FUNCTION "FRK_LineSetWalk" : Bool
{ S7_Optimized_Access := 'TRUE' }
VERSION : 0.1
VAR_INPUT
    RootIndex : Int;
    Scope : String;
    Phase : Int;
    Access : "FRK_Access";
    Ready : Bool;
END_VAR
VAR_TEMP
    Slot : Int;
END_VAR
BEGIN
    #FRK_LineSetWalk := FALSE;
    "FRK_SetRuntime".Work[#RootIndex].RejectScope := 'BenchLineOwner';
    IF NOT "FRK_LineScope"(Scope := #Scope) OR NOT "FRK_Line".Data.Applied
        OR "FRK_Line".Data.Status.Role <> 1 THEN RETURN; END_IF;
    IF #Phase = 2 THEN
        "FRK_Line".Data.Values := "FRK_LineSetStage".Values;
        "FRK_LineCommit"(State := "FRK_Line".Data);
        #FRK_LineSetWalk := TRUE; RETURN;
    END_IF;
    IF #Phase = 1 OR #Phase = 4 THEN "FRK_LineSetStage".Values := "FRK_Line".Data.Values; END_IF;
    "FRK_LineDef"(FieldIndex := 1);
    "FRK_SetRuntime".Work[#RootIndex].RejectScope := #Scope; "FRK_SetRuntime".Work[#RootIndex].RejectKey := "FRK_ConfigScratch".Entry.WriteKey;
    IF #Phase = 0 OR #Phase = 5 THEN
        IF #Phase = 5 AND NOT "FRK_ConfigDataAllowed"(Access := #Access, ForWrite := FALSE, Scope := #Scope) THEN RETURN; END_IF;
        "FRK_LineValue"(FieldIndex := 1, Values := "FRK_Line".Data.Values);
        IF NOT "FRK_ConfigValidate"(Text := "FRK_ConfigScratch".Entry.ValueText)
            OR "FRK_SetRuntime".Work[#RootIndex].Payload.Info.RecordCount >= 29 THEN RETURN; END_IF;
        #Slot := "FRK_SetRuntime".Work[#RootIndex].Payload.Info.RecordCount + 1;
        "FRK_SetRuntime".Work[#RootIndex].Payload.Records[#Slot].Scope := #Scope;
        "FRK_SetRuntime".Work[#RootIndex].Payload.Records[#Slot].WriteKey := "FRK_ConfigScratch".Entry.WriteKey;
        "FRK_SetRuntime".Work[#RootIndex].Payload.Records[#Slot].Revision := "FRK_ConfigScratch".Entry.WriteRevision;
        "FRK_SetRuntime".Work[#RootIndex].Payload.Records[#Slot].Kind := "FRK_ConfigScratch".Entry.ConfigKind;
        "FRK_SetRuntime".Work[#RootIndex].Payload.Records[#Slot].ValueType := "FRK_ConfigScratch".Entry.ValueType;
        "FRK_SetRuntime".Work[#RootIndex].Payload.Records[#Slot].ValueText := WSTRING_TO_STRING("FRK_ConfigScratch".Entry.ValueText);
        "FRK_SetRuntime".Work[#RootIndex].Payload.Info.RecordCount := #Slot;
    ELSE
        #Slot := "FRK_SetCheck"(RootIndex := #RootIndex, Scope := #Scope, Access := #Access, Ready := #Ready AND (#Phase = 4 OR "FRK_Line".Ready), WriteAccess := #Phase <> 3, ReserveTarget := FALSE);
        IF #Slot = 0 THEN RETURN; END_IF;
        IF #Phase = 1 OR #Phase = 4 THEN
    "FRK_LineSetStage".Values.TaktMs := LINT_TO_UDINT("FRK_ConfigScratch".Value.Number);
        END_IF;
    END_IF;
    "FRK_LineDef"(FieldIndex := 2);
    "FRK_SetRuntime".Work[#RootIndex].RejectScope := #Scope; "FRK_SetRuntime".Work[#RootIndex].RejectKey := "FRK_ConfigScratch".Entry.WriteKey;
    IF #Phase = 0 OR #Phase = 5 THEN
        IF #Phase = 5 AND NOT "FRK_ConfigDataAllowed"(Access := #Access, ForWrite := FALSE, Scope := #Scope) THEN RETURN; END_IF;
        "FRK_LineValue"(FieldIndex := 2, Values := "FRK_Line".Data.Values);
        IF NOT "FRK_ConfigValidate"(Text := "FRK_ConfigScratch".Entry.ValueText)
            OR "FRK_SetRuntime".Work[#RootIndex].Payload.Info.RecordCount >= 29 THEN RETURN; END_IF;
        #Slot := "FRK_SetRuntime".Work[#RootIndex].Payload.Info.RecordCount + 1;
        "FRK_SetRuntime".Work[#RootIndex].Payload.Records[#Slot].Scope := #Scope;
        "FRK_SetRuntime".Work[#RootIndex].Payload.Records[#Slot].WriteKey := "FRK_ConfigScratch".Entry.WriteKey;
        "FRK_SetRuntime".Work[#RootIndex].Payload.Records[#Slot].Revision := "FRK_ConfigScratch".Entry.WriteRevision;
        "FRK_SetRuntime".Work[#RootIndex].Payload.Records[#Slot].Kind := "FRK_ConfigScratch".Entry.ConfigKind;
        "FRK_SetRuntime".Work[#RootIndex].Payload.Records[#Slot].ValueType := "FRK_ConfigScratch".Entry.ValueType;
        "FRK_SetRuntime".Work[#RootIndex].Payload.Records[#Slot].ValueText := WSTRING_TO_STRING("FRK_ConfigScratch".Entry.ValueText);
        "FRK_SetRuntime".Work[#RootIndex].Payload.Info.RecordCount := #Slot;
    ELSE
        #Slot := "FRK_SetCheck"(RootIndex := #RootIndex, Scope := #Scope, Access := #Access, Ready := #Ready AND (#Phase = 4 OR "FRK_Line".Ready), WriteAccess := #Phase <> 3, ReserveTarget := FALSE);
        IF #Slot = 0 THEN RETURN; END_IF;
        IF #Phase = 1 OR #Phase = 4 THEN
    "FRK_LineSetStage".Values.Gain := "FRK_ConfigScratch".Value.Decimal;
        END_IF;
    END_IF;
    "FRK_LineDef"(FieldIndex := 3);
    "FRK_SetRuntime".Work[#RootIndex].RejectScope := #Scope; "FRK_SetRuntime".Work[#RootIndex].RejectKey := "FRK_ConfigScratch".Entry.WriteKey;
    IF #Phase = 0 OR #Phase = 5 THEN
        IF #Phase = 5 AND NOT "FRK_ConfigDataAllowed"(Access := #Access, ForWrite := FALSE, Scope := #Scope) THEN RETURN; END_IF;
        "FRK_LineValue"(FieldIndex := 3, Values := "FRK_Line".Data.Values);
        IF NOT "FRK_ConfigValidate"(Text := "FRK_ConfigScratch".Entry.ValueText)
            OR "FRK_SetRuntime".Work[#RootIndex].Payload.Info.RecordCount >= 29 THEN RETURN; END_IF;
        #Slot := "FRK_SetRuntime".Work[#RootIndex].Payload.Info.RecordCount + 1;
        "FRK_SetRuntime".Work[#RootIndex].Payload.Records[#Slot].Scope := #Scope;
        "FRK_SetRuntime".Work[#RootIndex].Payload.Records[#Slot].WriteKey := "FRK_ConfigScratch".Entry.WriteKey;
        "FRK_SetRuntime".Work[#RootIndex].Payload.Records[#Slot].Revision := "FRK_ConfigScratch".Entry.WriteRevision;
        "FRK_SetRuntime".Work[#RootIndex].Payload.Records[#Slot].Kind := "FRK_ConfigScratch".Entry.ConfigKind;
        "FRK_SetRuntime".Work[#RootIndex].Payload.Records[#Slot].ValueType := "FRK_ConfigScratch".Entry.ValueType;
        "FRK_SetRuntime".Work[#RootIndex].Payload.Records[#Slot].ValueText := WSTRING_TO_STRING("FRK_ConfigScratch".Entry.ValueText);
        "FRK_SetRuntime".Work[#RootIndex].Payload.Info.RecordCount := #Slot;
    ELSE
        #Slot := "FRK_SetCheck"(RootIndex := #RootIndex, Scope := #Scope, Access := #Access, Ready := #Ready AND (#Phase = 4 OR "FRK_Line".Ready), WriteAccess := #Phase <> 3, ReserveTarget := FALSE);
        IF #Slot = 0 THEN RETURN; END_IF;
        IF #Phase = 1 OR #Phase = 4 THEN
    "FRK_LineSetStage".Values.Grade := LINT_TO_DINT("FRK_ConfigScratch".Value.Number);
        END_IF;
    END_IF;
    "FRK_LineDef"(FieldIndex := 4);
    "FRK_SetRuntime".Work[#RootIndex].RejectScope := #Scope; "FRK_SetRuntime".Work[#RootIndex].RejectKey := "FRK_ConfigScratch".Entry.WriteKey;
    IF #Phase = 0 OR #Phase = 5 THEN
        IF #Phase = 5 AND NOT "FRK_ConfigDataAllowed"(Access := #Access, ForWrite := FALSE, Scope := #Scope) THEN RETURN; END_IF;
        "FRK_LineValue"(FieldIndex := 4, Values := "FRK_Line".Data.Values);
        IF NOT "FRK_ConfigValidate"(Text := "FRK_ConfigScratch".Entry.ValueText)
            OR "FRK_SetRuntime".Work[#RootIndex].Payload.Info.RecordCount >= 29 THEN RETURN; END_IF;
        #Slot := "FRK_SetRuntime".Work[#RootIndex].Payload.Info.RecordCount + 1;
        "FRK_SetRuntime".Work[#RootIndex].Payload.Records[#Slot].Scope := #Scope;
        "FRK_SetRuntime".Work[#RootIndex].Payload.Records[#Slot].WriteKey := "FRK_ConfigScratch".Entry.WriteKey;
        "FRK_SetRuntime".Work[#RootIndex].Payload.Records[#Slot].Revision := "FRK_ConfigScratch".Entry.WriteRevision;
        "FRK_SetRuntime".Work[#RootIndex].Payload.Records[#Slot].Kind := "FRK_ConfigScratch".Entry.ConfigKind;
        "FRK_SetRuntime".Work[#RootIndex].Payload.Records[#Slot].ValueType := "FRK_ConfigScratch".Entry.ValueType;
        "FRK_SetRuntime".Work[#RootIndex].Payload.Records[#Slot].ValueText := WSTRING_TO_STRING("FRK_ConfigScratch".Entry.ValueText);
        "FRK_SetRuntime".Work[#RootIndex].Payload.Info.RecordCount := #Slot;
    ELSE
        #Slot := "FRK_SetCheck"(RootIndex := #RootIndex, Scope := #Scope, Access := #Access, Ready := #Ready AND (#Phase = 4 OR "FRK_Line".Ready), WriteAccess := #Phase <> 3, ReserveTarget := FALSE);
        IF #Slot = 0 THEN RETURN; END_IF;
        IF #Phase = 1 OR #Phase = 4 THEN
    "FRK_LineSetStage".Values.Enabled := "FRK_ConfigScratch".Value.Flag;
        END_IF;
    END_IF;
    "FRK_LineDef"(FieldIndex := 5);
    "FRK_SetRuntime".Work[#RootIndex].RejectScope := #Scope; "FRK_SetRuntime".Work[#RootIndex].RejectKey := "FRK_ConfigScratch".Entry.WriteKey;
    IF #Phase = 0 OR #Phase = 5 THEN
        IF #Phase = 5 AND NOT "FRK_ConfigDataAllowed"(Access := #Access, ForWrite := FALSE, Scope := #Scope) THEN RETURN; END_IF;
        "FRK_LineValue"(FieldIndex := 5, Values := "FRK_Line".Data.Values);
        IF NOT "FRK_ConfigValidate"(Text := "FRK_ConfigScratch".Entry.ValueText)
            OR "FRK_SetRuntime".Work[#RootIndex].Payload.Info.RecordCount >= 29 THEN RETURN; END_IF;
        #Slot := "FRK_SetRuntime".Work[#RootIndex].Payload.Info.RecordCount + 1;
        "FRK_SetRuntime".Work[#RootIndex].Payload.Records[#Slot].Scope := #Scope;
        "FRK_SetRuntime".Work[#RootIndex].Payload.Records[#Slot].WriteKey := "FRK_ConfigScratch".Entry.WriteKey;
        "FRK_SetRuntime".Work[#RootIndex].Payload.Records[#Slot].Revision := "FRK_ConfigScratch".Entry.WriteRevision;
        "FRK_SetRuntime".Work[#RootIndex].Payload.Records[#Slot].Kind := "FRK_ConfigScratch".Entry.ConfigKind;
        "FRK_SetRuntime".Work[#RootIndex].Payload.Records[#Slot].ValueType := "FRK_ConfigScratch".Entry.ValueType;
        "FRK_SetRuntime".Work[#RootIndex].Payload.Records[#Slot].ValueText := WSTRING_TO_STRING("FRK_ConfigScratch".Entry.ValueText);
        "FRK_SetRuntime".Work[#RootIndex].Payload.Info.RecordCount := #Slot;
    ELSE
        #Slot := "FRK_SetCheck"(RootIndex := #RootIndex, Scope := #Scope, Access := #Access, Ready := #Ready AND (#Phase = 4 OR "FRK_Line".Ready), WriteAccess := #Phase <> 3, ReserveTarget := FALSE);
        IF #Slot = 0 THEN RETURN; END_IF;
        IF #Phase = 1 OR #Phase = 4 THEN
    "FRK_LineSetStage".Values.HostName := "FRK_ConfigScratch".Value.Text;
        END_IF;
    END_IF;
    "FRK_LineDef"(FieldIndex := 6);
    "FRK_SetRuntime".Work[#RootIndex].RejectScope := #Scope; "FRK_SetRuntime".Work[#RootIndex].RejectKey := "FRK_ConfigScratch".Entry.WriteKey;
    IF #Phase = 0 OR #Phase = 5 THEN
        IF #Phase = 5 AND NOT "FRK_ConfigDataAllowed"(Access := #Access, ForWrite := FALSE, Scope := #Scope) THEN RETURN; END_IF;
        "FRK_LineValue"(FieldIndex := 6, Values := "FRK_Line".Data.Values);
        IF NOT "FRK_ConfigValidate"(Text := "FRK_ConfigScratch".Entry.ValueText)
            OR "FRK_SetRuntime".Work[#RootIndex].Payload.Info.RecordCount >= 29 THEN RETURN; END_IF;
        #Slot := "FRK_SetRuntime".Work[#RootIndex].Payload.Info.RecordCount + 1;
        "FRK_SetRuntime".Work[#RootIndex].Payload.Records[#Slot].Scope := #Scope;
        "FRK_SetRuntime".Work[#RootIndex].Payload.Records[#Slot].WriteKey := "FRK_ConfigScratch".Entry.WriteKey;
        "FRK_SetRuntime".Work[#RootIndex].Payload.Records[#Slot].Revision := "FRK_ConfigScratch".Entry.WriteRevision;
        "FRK_SetRuntime".Work[#RootIndex].Payload.Records[#Slot].Kind := "FRK_ConfigScratch".Entry.ConfigKind;
        "FRK_SetRuntime".Work[#RootIndex].Payload.Records[#Slot].ValueType := "FRK_ConfigScratch".Entry.ValueType;
        "FRK_SetRuntime".Work[#RootIndex].Payload.Records[#Slot].ValueText := WSTRING_TO_STRING("FRK_ConfigScratch".Entry.ValueText);
        "FRK_SetRuntime".Work[#RootIndex].Payload.Info.RecordCount := #Slot;
    ELSE
        #Slot := "FRK_SetCheck"(RootIndex := #RootIndex, Scope := #Scope, Access := #Access, Ready := #Ready AND (#Phase = 4 OR "FRK_Line".Ready), WriteAccess := #Phase <> 3, ReserveTarget := FALSE);
        IF #Slot = 0 THEN RETURN; END_IF;
        IF #Phase = 1 OR #Phase = 4 THEN
    "FRK_LineSetStage".Values.Offsets[0] := LINT_TO_INT("FRK_ConfigScratch".Value.Number);
        END_IF;
    END_IF;
    "FRK_LineDef"(FieldIndex := 7);
    "FRK_SetRuntime".Work[#RootIndex].RejectScope := #Scope; "FRK_SetRuntime".Work[#RootIndex].RejectKey := "FRK_ConfigScratch".Entry.WriteKey;
    IF #Phase = 0 OR #Phase = 5 THEN
        IF #Phase = 5 AND NOT "FRK_ConfigDataAllowed"(Access := #Access, ForWrite := FALSE, Scope := #Scope) THEN RETURN; END_IF;
        "FRK_LineValue"(FieldIndex := 7, Values := "FRK_Line".Data.Values);
        IF NOT "FRK_ConfigValidate"(Text := "FRK_ConfigScratch".Entry.ValueText)
            OR "FRK_SetRuntime".Work[#RootIndex].Payload.Info.RecordCount >= 29 THEN RETURN; END_IF;
        #Slot := "FRK_SetRuntime".Work[#RootIndex].Payload.Info.RecordCount + 1;
        "FRK_SetRuntime".Work[#RootIndex].Payload.Records[#Slot].Scope := #Scope;
        "FRK_SetRuntime".Work[#RootIndex].Payload.Records[#Slot].WriteKey := "FRK_ConfigScratch".Entry.WriteKey;
        "FRK_SetRuntime".Work[#RootIndex].Payload.Records[#Slot].Revision := "FRK_ConfigScratch".Entry.WriteRevision;
        "FRK_SetRuntime".Work[#RootIndex].Payload.Records[#Slot].Kind := "FRK_ConfigScratch".Entry.ConfigKind;
        "FRK_SetRuntime".Work[#RootIndex].Payload.Records[#Slot].ValueType := "FRK_ConfigScratch".Entry.ValueType;
        "FRK_SetRuntime".Work[#RootIndex].Payload.Records[#Slot].ValueText := WSTRING_TO_STRING("FRK_ConfigScratch".Entry.ValueText);
        "FRK_SetRuntime".Work[#RootIndex].Payload.Info.RecordCount := #Slot;
    ELSE
        #Slot := "FRK_SetCheck"(RootIndex := #RootIndex, Scope := #Scope, Access := #Access, Ready := #Ready AND (#Phase = 4 OR "FRK_Line".Ready), WriteAccess := #Phase <> 3, ReserveTarget := FALSE);
        IF #Slot = 0 THEN RETURN; END_IF;
        IF #Phase = 1 OR #Phase = 4 THEN
    "FRK_LineSetStage".Values.Offsets[1] := LINT_TO_INT("FRK_ConfigScratch".Value.Number);
        END_IF;
    END_IF;
    "FRK_LineDef"(FieldIndex := 8);
    "FRK_SetRuntime".Work[#RootIndex].RejectScope := #Scope; "FRK_SetRuntime".Work[#RootIndex].RejectKey := "FRK_ConfigScratch".Entry.WriteKey;
    IF #Phase = 0 OR #Phase = 5 THEN
        IF #Phase = 5 AND NOT "FRK_ConfigDataAllowed"(Access := #Access, ForWrite := FALSE, Scope := #Scope) THEN RETURN; END_IF;
        "FRK_LineValue"(FieldIndex := 8, Values := "FRK_Line".Data.Values);
        IF NOT "FRK_ConfigValidate"(Text := "FRK_ConfigScratch".Entry.ValueText)
            OR "FRK_SetRuntime".Work[#RootIndex].Payload.Info.RecordCount >= 29 THEN RETURN; END_IF;
        #Slot := "FRK_SetRuntime".Work[#RootIndex].Payload.Info.RecordCount + 1;
        "FRK_SetRuntime".Work[#RootIndex].Payload.Records[#Slot].Scope := #Scope;
        "FRK_SetRuntime".Work[#RootIndex].Payload.Records[#Slot].WriteKey := "FRK_ConfigScratch".Entry.WriteKey;
        "FRK_SetRuntime".Work[#RootIndex].Payload.Records[#Slot].Revision := "FRK_ConfigScratch".Entry.WriteRevision;
        "FRK_SetRuntime".Work[#RootIndex].Payload.Records[#Slot].Kind := "FRK_ConfigScratch".Entry.ConfigKind;
        "FRK_SetRuntime".Work[#RootIndex].Payload.Records[#Slot].ValueType := "FRK_ConfigScratch".Entry.ValueType;
        "FRK_SetRuntime".Work[#RootIndex].Payload.Records[#Slot].ValueText := WSTRING_TO_STRING("FRK_ConfigScratch".Entry.ValueText);
        "FRK_SetRuntime".Work[#RootIndex].Payload.Info.RecordCount := #Slot;
    ELSE
        #Slot := "FRK_SetCheck"(RootIndex := #RootIndex, Scope := #Scope, Access := #Access, Ready := #Ready AND (#Phase = 4 OR "FRK_Line".Ready), WriteAccess := #Phase <> 3, ReserveTarget := FALSE);
        IF #Slot = 0 THEN RETURN; END_IF;
        IF #Phase = 1 OR #Phase = 4 THEN
    "FRK_LineSetStage".Values.Small := LINT_TO_USINT("FRK_ConfigScratch".Value.Number);
        END_IF;
    END_IF;
    "FRK_LineDef"(FieldIndex := 9);
    "FRK_SetRuntime".Work[#RootIndex].RejectScope := #Scope; "FRK_SetRuntime".Work[#RootIndex].RejectKey := "FRK_ConfigScratch".Entry.WriteKey;
    IF #Phase = 0 OR #Phase = 5 THEN
        IF #Phase = 5 AND NOT "FRK_ConfigDataAllowed"(Access := #Access, ForWrite := FALSE, Scope := #Scope) THEN RETURN; END_IF;
        "FRK_LineValue"(FieldIndex := 9, Values := "FRK_Line".Data.Values);
        IF NOT "FRK_ConfigValidate"(Text := "FRK_ConfigScratch".Entry.ValueText)
            OR "FRK_SetRuntime".Work[#RootIndex].Payload.Info.RecordCount >= 29 THEN RETURN; END_IF;
        #Slot := "FRK_SetRuntime".Work[#RootIndex].Payload.Info.RecordCount + 1;
        "FRK_SetRuntime".Work[#RootIndex].Payload.Records[#Slot].Scope := #Scope;
        "FRK_SetRuntime".Work[#RootIndex].Payload.Records[#Slot].WriteKey := "FRK_ConfigScratch".Entry.WriteKey;
        "FRK_SetRuntime".Work[#RootIndex].Payload.Records[#Slot].Revision := "FRK_ConfigScratch".Entry.WriteRevision;
        "FRK_SetRuntime".Work[#RootIndex].Payload.Records[#Slot].Kind := "FRK_ConfigScratch".Entry.ConfigKind;
        "FRK_SetRuntime".Work[#RootIndex].Payload.Records[#Slot].ValueType := "FRK_ConfigScratch".Entry.ValueType;
        "FRK_SetRuntime".Work[#RootIndex].Payload.Records[#Slot].ValueText := WSTRING_TO_STRING("FRK_ConfigScratch".Entry.ValueText);
        "FRK_SetRuntime".Work[#RootIndex].Payload.Info.RecordCount := #Slot;
    ELSE
        #Slot := "FRK_SetCheck"(RootIndex := #RootIndex, Scope := #Scope, Access := #Access, Ready := #Ready AND (#Phase = 4 OR "FRK_Line".Ready), WriteAccess := #Phase <> 3, ReserveTarget := FALSE);
        IF #Slot = 0 THEN RETURN; END_IF;
        IF #Phase = 1 OR #Phase = 4 THEN
    "FRK_LineSetStage".Values.UtcOffsetMin := LINT_TO_DINT("FRK_ConfigScratch".Value.Number);
        END_IF;
    END_IF;
    "FRK_LineDef"(FieldIndex := 10);
    "FRK_SetRuntime".Work[#RootIndex].RejectScope := #Scope; "FRK_SetRuntime".Work[#RootIndex].RejectKey := "FRK_ConfigScratch".Entry.WriteKey;
    IF #Phase = 0 OR #Phase = 5 THEN
        IF #Phase = 5 AND NOT "FRK_ConfigDataAllowed"(Access := #Access, ForWrite := FALSE, Scope := #Scope) THEN RETURN; END_IF;
        "FRK_LineValue"(FieldIndex := 10, Values := "FRK_Line".Data.Values);
        IF NOT "FRK_ConfigValidate"(Text := "FRK_ConfigScratch".Entry.ValueText)
            OR "FRK_SetRuntime".Work[#RootIndex].Payload.Info.RecordCount >= 29 THEN RETURN; END_IF;
        #Slot := "FRK_SetRuntime".Work[#RootIndex].Payload.Info.RecordCount + 1;
        "FRK_SetRuntime".Work[#RootIndex].Payload.Records[#Slot].Scope := #Scope;
        "FRK_SetRuntime".Work[#RootIndex].Payload.Records[#Slot].WriteKey := "FRK_ConfigScratch".Entry.WriteKey;
        "FRK_SetRuntime".Work[#RootIndex].Payload.Records[#Slot].Revision := "FRK_ConfigScratch".Entry.WriteRevision;
        "FRK_SetRuntime".Work[#RootIndex].Payload.Records[#Slot].Kind := "FRK_ConfigScratch".Entry.ConfigKind;
        "FRK_SetRuntime".Work[#RootIndex].Payload.Records[#Slot].ValueType := "FRK_ConfigScratch".Entry.ValueType;
        "FRK_SetRuntime".Work[#RootIndex].Payload.Records[#Slot].ValueText := WSTRING_TO_STRING("FRK_ConfigScratch".Entry.ValueText);
        "FRK_SetRuntime".Work[#RootIndex].Payload.Info.RecordCount := #Slot;
    ELSE
        #Slot := "FRK_SetCheck"(RootIndex := #RootIndex, Scope := #Scope, Access := #Access, Ready := #Ready AND (#Phase = 4 OR "FRK_Line".Ready), WriteAccess := #Phase <> 3, ReserveTarget := FALSE);
        IF #Slot = 0 THEN RETURN; END_IF;
        IF #Phase = 1 OR #Phase = 4 THEN
    "FRK_LineSetStage".Values.ShiftStartMin[1] := LINT_TO_DINT("FRK_ConfigScratch".Value.Number);
        END_IF;
    END_IF;
    "FRK_LineDef"(FieldIndex := 11);
    "FRK_SetRuntime".Work[#RootIndex].RejectScope := #Scope; "FRK_SetRuntime".Work[#RootIndex].RejectKey := "FRK_ConfigScratch".Entry.WriteKey;
    IF #Phase = 0 OR #Phase = 5 THEN
        IF #Phase = 5 AND NOT "FRK_ConfigDataAllowed"(Access := #Access, ForWrite := FALSE, Scope := #Scope) THEN RETURN; END_IF;
        "FRK_LineValue"(FieldIndex := 11, Values := "FRK_Line".Data.Values);
        IF NOT "FRK_ConfigValidate"(Text := "FRK_ConfigScratch".Entry.ValueText)
            OR "FRK_SetRuntime".Work[#RootIndex].Payload.Info.RecordCount >= 29 THEN RETURN; END_IF;
        #Slot := "FRK_SetRuntime".Work[#RootIndex].Payload.Info.RecordCount + 1;
        "FRK_SetRuntime".Work[#RootIndex].Payload.Records[#Slot].Scope := #Scope;
        "FRK_SetRuntime".Work[#RootIndex].Payload.Records[#Slot].WriteKey := "FRK_ConfigScratch".Entry.WriteKey;
        "FRK_SetRuntime".Work[#RootIndex].Payload.Records[#Slot].Revision := "FRK_ConfigScratch".Entry.WriteRevision;
        "FRK_SetRuntime".Work[#RootIndex].Payload.Records[#Slot].Kind := "FRK_ConfigScratch".Entry.ConfigKind;
        "FRK_SetRuntime".Work[#RootIndex].Payload.Records[#Slot].ValueType := "FRK_ConfigScratch".Entry.ValueType;
        "FRK_SetRuntime".Work[#RootIndex].Payload.Records[#Slot].ValueText := WSTRING_TO_STRING("FRK_ConfigScratch".Entry.ValueText);
        "FRK_SetRuntime".Work[#RootIndex].Payload.Info.RecordCount := #Slot;
    ELSE
        #Slot := "FRK_SetCheck"(RootIndex := #RootIndex, Scope := #Scope, Access := #Access, Ready := #Ready AND (#Phase = 4 OR "FRK_Line".Ready), WriteAccess := #Phase <> 3, ReserveTarget := FALSE);
        IF #Slot = 0 THEN RETURN; END_IF;
        IF #Phase = 1 OR #Phase = 4 THEN
    "FRK_LineSetStage".Values.ShiftDurationMin[1] := LINT_TO_DINT("FRK_ConfigScratch".Value.Number);
        END_IF;
    END_IF;
    "FRK_LineDef"(FieldIndex := 12);
    "FRK_SetRuntime".Work[#RootIndex].RejectScope := #Scope; "FRK_SetRuntime".Work[#RootIndex].RejectKey := "FRK_ConfigScratch".Entry.WriteKey;
    IF #Phase = 0 OR #Phase = 5 THEN
        IF #Phase = 5 AND NOT "FRK_ConfigDataAllowed"(Access := #Access, ForWrite := FALSE, Scope := #Scope) THEN RETURN; END_IF;
        "FRK_LineValue"(FieldIndex := 12, Values := "FRK_Line".Data.Values);
        IF NOT "FRK_ConfigValidate"(Text := "FRK_ConfigScratch".Entry.ValueText)
            OR "FRK_SetRuntime".Work[#RootIndex].Payload.Info.RecordCount >= 29 THEN RETURN; END_IF;
        #Slot := "FRK_SetRuntime".Work[#RootIndex].Payload.Info.RecordCount + 1;
        "FRK_SetRuntime".Work[#RootIndex].Payload.Records[#Slot].Scope := #Scope;
        "FRK_SetRuntime".Work[#RootIndex].Payload.Records[#Slot].WriteKey := "FRK_ConfigScratch".Entry.WriteKey;
        "FRK_SetRuntime".Work[#RootIndex].Payload.Records[#Slot].Revision := "FRK_ConfigScratch".Entry.WriteRevision;
        "FRK_SetRuntime".Work[#RootIndex].Payload.Records[#Slot].Kind := "FRK_ConfigScratch".Entry.ConfigKind;
        "FRK_SetRuntime".Work[#RootIndex].Payload.Records[#Slot].ValueType := "FRK_ConfigScratch".Entry.ValueType;
        "FRK_SetRuntime".Work[#RootIndex].Payload.Records[#Slot].ValueText := WSTRING_TO_STRING("FRK_ConfigScratch".Entry.ValueText);
        "FRK_SetRuntime".Work[#RootIndex].Payload.Info.RecordCount := #Slot;
    ELSE
        #Slot := "FRK_SetCheck"(RootIndex := #RootIndex, Scope := #Scope, Access := #Access, Ready := #Ready AND (#Phase = 4 OR "FRK_Line".Ready), WriteAccess := #Phase <> 3, ReserveTarget := FALSE);
        IF #Slot = 0 THEN RETURN; END_IF;
        IF #Phase = 1 OR #Phase = 4 THEN
    "FRK_LineSetStage".Values.ShiftActiveDays[1] := LINT_TO_DINT("FRK_ConfigScratch".Value.Number);
        END_IF;
    END_IF;
    "FRK_LineDef"(FieldIndex := 13);
    "FRK_SetRuntime".Work[#RootIndex].RejectScope := #Scope; "FRK_SetRuntime".Work[#RootIndex].RejectKey := "FRK_ConfigScratch".Entry.WriteKey;
    IF #Phase = 0 OR #Phase = 5 THEN
        IF #Phase = 5 AND NOT "FRK_ConfigDataAllowed"(Access := #Access, ForWrite := FALSE, Scope := #Scope) THEN RETURN; END_IF;
        "FRK_LineValue"(FieldIndex := 13, Values := "FRK_Line".Data.Values);
        IF NOT "FRK_ConfigValidate"(Text := "FRK_ConfigScratch".Entry.ValueText)
            OR "FRK_SetRuntime".Work[#RootIndex].Payload.Info.RecordCount >= 29 THEN RETURN; END_IF;
        #Slot := "FRK_SetRuntime".Work[#RootIndex].Payload.Info.RecordCount + 1;
        "FRK_SetRuntime".Work[#RootIndex].Payload.Records[#Slot].Scope := #Scope;
        "FRK_SetRuntime".Work[#RootIndex].Payload.Records[#Slot].WriteKey := "FRK_ConfigScratch".Entry.WriteKey;
        "FRK_SetRuntime".Work[#RootIndex].Payload.Records[#Slot].Revision := "FRK_ConfigScratch".Entry.WriteRevision;
        "FRK_SetRuntime".Work[#RootIndex].Payload.Records[#Slot].Kind := "FRK_ConfigScratch".Entry.ConfigKind;
        "FRK_SetRuntime".Work[#RootIndex].Payload.Records[#Slot].ValueType := "FRK_ConfigScratch".Entry.ValueType;
        "FRK_SetRuntime".Work[#RootIndex].Payload.Records[#Slot].ValueText := WSTRING_TO_STRING("FRK_ConfigScratch".Entry.ValueText);
        "FRK_SetRuntime".Work[#RootIndex].Payload.Info.RecordCount := #Slot;
    ELSE
        #Slot := "FRK_SetCheck"(RootIndex := #RootIndex, Scope := #Scope, Access := #Access, Ready := #Ready AND (#Phase = 4 OR "FRK_Line".Ready), WriteAccess := #Phase <> 3, ReserveTarget := FALSE);
        IF #Slot = 0 THEN RETURN; END_IF;
        IF #Phase = 1 OR #Phase = 4 THEN
    "FRK_LineSetStage".Values.ShiftTarget[1] := LINT_TO_DINT("FRK_ConfigScratch".Value.Number);
        END_IF;
    END_IF;
    "FRK_LineDef"(FieldIndex := 14);
    "FRK_SetRuntime".Work[#RootIndex].RejectScope := #Scope; "FRK_SetRuntime".Work[#RootIndex].RejectKey := "FRK_ConfigScratch".Entry.WriteKey;
    IF #Phase = 0 OR #Phase = 5 THEN
        IF #Phase = 5 AND NOT "FRK_ConfigDataAllowed"(Access := #Access, ForWrite := FALSE, Scope := #Scope) THEN RETURN; END_IF;
        "FRK_LineValue"(FieldIndex := 14, Values := "FRK_Line".Data.Values);
        IF NOT "FRK_ConfigValidate"(Text := "FRK_ConfigScratch".Entry.ValueText)
            OR "FRK_SetRuntime".Work[#RootIndex].Payload.Info.RecordCount >= 29 THEN RETURN; END_IF;
        #Slot := "FRK_SetRuntime".Work[#RootIndex].Payload.Info.RecordCount + 1;
        "FRK_SetRuntime".Work[#RootIndex].Payload.Records[#Slot].Scope := #Scope;
        "FRK_SetRuntime".Work[#RootIndex].Payload.Records[#Slot].WriteKey := "FRK_ConfigScratch".Entry.WriteKey;
        "FRK_SetRuntime".Work[#RootIndex].Payload.Records[#Slot].Revision := "FRK_ConfigScratch".Entry.WriteRevision;
        "FRK_SetRuntime".Work[#RootIndex].Payload.Records[#Slot].Kind := "FRK_ConfigScratch".Entry.ConfigKind;
        "FRK_SetRuntime".Work[#RootIndex].Payload.Records[#Slot].ValueType := "FRK_ConfigScratch".Entry.ValueType;
        "FRK_SetRuntime".Work[#RootIndex].Payload.Records[#Slot].ValueText := WSTRING_TO_STRING("FRK_ConfigScratch".Entry.ValueText);
        "FRK_SetRuntime".Work[#RootIndex].Payload.Info.RecordCount := #Slot;
    ELSE
        #Slot := "FRK_SetCheck"(RootIndex := #RootIndex, Scope := #Scope, Access := #Access, Ready := #Ready AND (#Phase = 4 OR "FRK_Line".Ready), WriteAccess := #Phase <> 3, ReserveTarget := FALSE);
        IF #Slot = 0 THEN RETURN; END_IF;
        IF #Phase = 1 OR #Phase = 4 THEN
    "FRK_LineSetStage".Values.ShiftStartMin[2] := LINT_TO_DINT("FRK_ConfigScratch".Value.Number);
        END_IF;
    END_IF;
    "FRK_LineDef"(FieldIndex := 15);
    "FRK_SetRuntime".Work[#RootIndex].RejectScope := #Scope; "FRK_SetRuntime".Work[#RootIndex].RejectKey := "FRK_ConfigScratch".Entry.WriteKey;
    IF #Phase = 0 OR #Phase = 5 THEN
        IF #Phase = 5 AND NOT "FRK_ConfigDataAllowed"(Access := #Access, ForWrite := FALSE, Scope := #Scope) THEN RETURN; END_IF;
        "FRK_LineValue"(FieldIndex := 15, Values := "FRK_Line".Data.Values);
        IF NOT "FRK_ConfigValidate"(Text := "FRK_ConfigScratch".Entry.ValueText)
            OR "FRK_SetRuntime".Work[#RootIndex].Payload.Info.RecordCount >= 29 THEN RETURN; END_IF;
        #Slot := "FRK_SetRuntime".Work[#RootIndex].Payload.Info.RecordCount + 1;
        "FRK_SetRuntime".Work[#RootIndex].Payload.Records[#Slot].Scope := #Scope;
        "FRK_SetRuntime".Work[#RootIndex].Payload.Records[#Slot].WriteKey := "FRK_ConfigScratch".Entry.WriteKey;
        "FRK_SetRuntime".Work[#RootIndex].Payload.Records[#Slot].Revision := "FRK_ConfigScratch".Entry.WriteRevision;
        "FRK_SetRuntime".Work[#RootIndex].Payload.Records[#Slot].Kind := "FRK_ConfigScratch".Entry.ConfigKind;
        "FRK_SetRuntime".Work[#RootIndex].Payload.Records[#Slot].ValueType := "FRK_ConfigScratch".Entry.ValueType;
        "FRK_SetRuntime".Work[#RootIndex].Payload.Records[#Slot].ValueText := WSTRING_TO_STRING("FRK_ConfigScratch".Entry.ValueText);
        "FRK_SetRuntime".Work[#RootIndex].Payload.Info.RecordCount := #Slot;
    ELSE
        #Slot := "FRK_SetCheck"(RootIndex := #RootIndex, Scope := #Scope, Access := #Access, Ready := #Ready AND (#Phase = 4 OR "FRK_Line".Ready), WriteAccess := #Phase <> 3, ReserveTarget := FALSE);
        IF #Slot = 0 THEN RETURN; END_IF;
        IF #Phase = 1 OR #Phase = 4 THEN
    "FRK_LineSetStage".Values.ShiftDurationMin[2] := LINT_TO_DINT("FRK_ConfigScratch".Value.Number);
        END_IF;
    END_IF;
    "FRK_LineDef"(FieldIndex := 16);
    "FRK_SetRuntime".Work[#RootIndex].RejectScope := #Scope; "FRK_SetRuntime".Work[#RootIndex].RejectKey := "FRK_ConfigScratch".Entry.WriteKey;
    IF #Phase = 0 OR #Phase = 5 THEN
        IF #Phase = 5 AND NOT "FRK_ConfigDataAllowed"(Access := #Access, ForWrite := FALSE, Scope := #Scope) THEN RETURN; END_IF;
        "FRK_LineValue"(FieldIndex := 16, Values := "FRK_Line".Data.Values);
        IF NOT "FRK_ConfigValidate"(Text := "FRK_ConfigScratch".Entry.ValueText)
            OR "FRK_SetRuntime".Work[#RootIndex].Payload.Info.RecordCount >= 29 THEN RETURN; END_IF;
        #Slot := "FRK_SetRuntime".Work[#RootIndex].Payload.Info.RecordCount + 1;
        "FRK_SetRuntime".Work[#RootIndex].Payload.Records[#Slot].Scope := #Scope;
        "FRK_SetRuntime".Work[#RootIndex].Payload.Records[#Slot].WriteKey := "FRK_ConfigScratch".Entry.WriteKey;
        "FRK_SetRuntime".Work[#RootIndex].Payload.Records[#Slot].Revision := "FRK_ConfigScratch".Entry.WriteRevision;
        "FRK_SetRuntime".Work[#RootIndex].Payload.Records[#Slot].Kind := "FRK_ConfigScratch".Entry.ConfigKind;
        "FRK_SetRuntime".Work[#RootIndex].Payload.Records[#Slot].ValueType := "FRK_ConfigScratch".Entry.ValueType;
        "FRK_SetRuntime".Work[#RootIndex].Payload.Records[#Slot].ValueText := WSTRING_TO_STRING("FRK_ConfigScratch".Entry.ValueText);
        "FRK_SetRuntime".Work[#RootIndex].Payload.Info.RecordCount := #Slot;
    ELSE
        #Slot := "FRK_SetCheck"(RootIndex := #RootIndex, Scope := #Scope, Access := #Access, Ready := #Ready AND (#Phase = 4 OR "FRK_Line".Ready), WriteAccess := #Phase <> 3, ReserveTarget := FALSE);
        IF #Slot = 0 THEN RETURN; END_IF;
        IF #Phase = 1 OR #Phase = 4 THEN
    "FRK_LineSetStage".Values.ShiftActiveDays[2] := LINT_TO_DINT("FRK_ConfigScratch".Value.Number);
        END_IF;
    END_IF;
    "FRK_LineDef"(FieldIndex := 17);
    "FRK_SetRuntime".Work[#RootIndex].RejectScope := #Scope; "FRK_SetRuntime".Work[#RootIndex].RejectKey := "FRK_ConfigScratch".Entry.WriteKey;
    IF #Phase = 0 OR #Phase = 5 THEN
        IF #Phase = 5 AND NOT "FRK_ConfigDataAllowed"(Access := #Access, ForWrite := FALSE, Scope := #Scope) THEN RETURN; END_IF;
        "FRK_LineValue"(FieldIndex := 17, Values := "FRK_Line".Data.Values);
        IF NOT "FRK_ConfigValidate"(Text := "FRK_ConfigScratch".Entry.ValueText)
            OR "FRK_SetRuntime".Work[#RootIndex].Payload.Info.RecordCount >= 29 THEN RETURN; END_IF;
        #Slot := "FRK_SetRuntime".Work[#RootIndex].Payload.Info.RecordCount + 1;
        "FRK_SetRuntime".Work[#RootIndex].Payload.Records[#Slot].Scope := #Scope;
        "FRK_SetRuntime".Work[#RootIndex].Payload.Records[#Slot].WriteKey := "FRK_ConfigScratch".Entry.WriteKey;
        "FRK_SetRuntime".Work[#RootIndex].Payload.Records[#Slot].Revision := "FRK_ConfigScratch".Entry.WriteRevision;
        "FRK_SetRuntime".Work[#RootIndex].Payload.Records[#Slot].Kind := "FRK_ConfigScratch".Entry.ConfigKind;
        "FRK_SetRuntime".Work[#RootIndex].Payload.Records[#Slot].ValueType := "FRK_ConfigScratch".Entry.ValueType;
        "FRK_SetRuntime".Work[#RootIndex].Payload.Records[#Slot].ValueText := WSTRING_TO_STRING("FRK_ConfigScratch".Entry.ValueText);
        "FRK_SetRuntime".Work[#RootIndex].Payload.Info.RecordCount := #Slot;
    ELSE
        #Slot := "FRK_SetCheck"(RootIndex := #RootIndex, Scope := #Scope, Access := #Access, Ready := #Ready AND (#Phase = 4 OR "FRK_Line".Ready), WriteAccess := #Phase <> 3, ReserveTarget := FALSE);
        IF #Slot = 0 THEN RETURN; END_IF;
        IF #Phase = 1 OR #Phase = 4 THEN
    "FRK_LineSetStage".Values.ShiftTarget[2] := LINT_TO_DINT("FRK_ConfigScratch".Value.Number);
        END_IF;
    END_IF;
    "FRK_LineDef"(FieldIndex := 18);
    "FRK_SetRuntime".Work[#RootIndex].RejectScope := #Scope; "FRK_SetRuntime".Work[#RootIndex].RejectKey := "FRK_ConfigScratch".Entry.WriteKey;
    IF #Phase = 0 OR #Phase = 5 THEN
        IF #Phase = 5 AND NOT "FRK_ConfigDataAllowed"(Access := #Access, ForWrite := FALSE, Scope := #Scope) THEN RETURN; END_IF;
        "FRK_LineValue"(FieldIndex := 18, Values := "FRK_Line".Data.Values);
        IF NOT "FRK_ConfigValidate"(Text := "FRK_ConfigScratch".Entry.ValueText)
            OR "FRK_SetRuntime".Work[#RootIndex].Payload.Info.RecordCount >= 29 THEN RETURN; END_IF;
        #Slot := "FRK_SetRuntime".Work[#RootIndex].Payload.Info.RecordCount + 1;
        "FRK_SetRuntime".Work[#RootIndex].Payload.Records[#Slot].Scope := #Scope;
        "FRK_SetRuntime".Work[#RootIndex].Payload.Records[#Slot].WriteKey := "FRK_ConfigScratch".Entry.WriteKey;
        "FRK_SetRuntime".Work[#RootIndex].Payload.Records[#Slot].Revision := "FRK_ConfigScratch".Entry.WriteRevision;
        "FRK_SetRuntime".Work[#RootIndex].Payload.Records[#Slot].Kind := "FRK_ConfigScratch".Entry.ConfigKind;
        "FRK_SetRuntime".Work[#RootIndex].Payload.Records[#Slot].ValueType := "FRK_ConfigScratch".Entry.ValueType;
        "FRK_SetRuntime".Work[#RootIndex].Payload.Records[#Slot].ValueText := WSTRING_TO_STRING("FRK_ConfigScratch".Entry.ValueText);
        "FRK_SetRuntime".Work[#RootIndex].Payload.Info.RecordCount := #Slot;
    ELSE
        #Slot := "FRK_SetCheck"(RootIndex := #RootIndex, Scope := #Scope, Access := #Access, Ready := #Ready AND (#Phase = 4 OR "FRK_Line".Ready), WriteAccess := #Phase <> 3, ReserveTarget := FALSE);
        IF #Slot = 0 THEN RETURN; END_IF;
        IF #Phase = 1 OR #Phase = 4 THEN
    "FRK_LineSetStage".Values.ShiftStartMin[3] := LINT_TO_DINT("FRK_ConfigScratch".Value.Number);
        END_IF;
    END_IF;
    "FRK_LineDef"(FieldIndex := 19);
    "FRK_SetRuntime".Work[#RootIndex].RejectScope := #Scope; "FRK_SetRuntime".Work[#RootIndex].RejectKey := "FRK_ConfigScratch".Entry.WriteKey;
    IF #Phase = 0 OR #Phase = 5 THEN
        IF #Phase = 5 AND NOT "FRK_ConfigDataAllowed"(Access := #Access, ForWrite := FALSE, Scope := #Scope) THEN RETURN; END_IF;
        "FRK_LineValue"(FieldIndex := 19, Values := "FRK_Line".Data.Values);
        IF NOT "FRK_ConfigValidate"(Text := "FRK_ConfigScratch".Entry.ValueText)
            OR "FRK_SetRuntime".Work[#RootIndex].Payload.Info.RecordCount >= 29 THEN RETURN; END_IF;
        #Slot := "FRK_SetRuntime".Work[#RootIndex].Payload.Info.RecordCount + 1;
        "FRK_SetRuntime".Work[#RootIndex].Payload.Records[#Slot].Scope := #Scope;
        "FRK_SetRuntime".Work[#RootIndex].Payload.Records[#Slot].WriteKey := "FRK_ConfigScratch".Entry.WriteKey;
        "FRK_SetRuntime".Work[#RootIndex].Payload.Records[#Slot].Revision := "FRK_ConfigScratch".Entry.WriteRevision;
        "FRK_SetRuntime".Work[#RootIndex].Payload.Records[#Slot].Kind := "FRK_ConfigScratch".Entry.ConfigKind;
        "FRK_SetRuntime".Work[#RootIndex].Payload.Records[#Slot].ValueType := "FRK_ConfigScratch".Entry.ValueType;
        "FRK_SetRuntime".Work[#RootIndex].Payload.Records[#Slot].ValueText := WSTRING_TO_STRING("FRK_ConfigScratch".Entry.ValueText);
        "FRK_SetRuntime".Work[#RootIndex].Payload.Info.RecordCount := #Slot;
    ELSE
        #Slot := "FRK_SetCheck"(RootIndex := #RootIndex, Scope := #Scope, Access := #Access, Ready := #Ready AND (#Phase = 4 OR "FRK_Line".Ready), WriteAccess := #Phase <> 3, ReserveTarget := FALSE);
        IF #Slot = 0 THEN RETURN; END_IF;
        IF #Phase = 1 OR #Phase = 4 THEN
    "FRK_LineSetStage".Values.ShiftDurationMin[3] := LINT_TO_DINT("FRK_ConfigScratch".Value.Number);
        END_IF;
    END_IF;
    "FRK_LineDef"(FieldIndex := 20);
    "FRK_SetRuntime".Work[#RootIndex].RejectScope := #Scope; "FRK_SetRuntime".Work[#RootIndex].RejectKey := "FRK_ConfigScratch".Entry.WriteKey;
    IF #Phase = 0 OR #Phase = 5 THEN
        IF #Phase = 5 AND NOT "FRK_ConfigDataAllowed"(Access := #Access, ForWrite := FALSE, Scope := #Scope) THEN RETURN; END_IF;
        "FRK_LineValue"(FieldIndex := 20, Values := "FRK_Line".Data.Values);
        IF NOT "FRK_ConfigValidate"(Text := "FRK_ConfigScratch".Entry.ValueText)
            OR "FRK_SetRuntime".Work[#RootIndex].Payload.Info.RecordCount >= 29 THEN RETURN; END_IF;
        #Slot := "FRK_SetRuntime".Work[#RootIndex].Payload.Info.RecordCount + 1;
        "FRK_SetRuntime".Work[#RootIndex].Payload.Records[#Slot].Scope := #Scope;
        "FRK_SetRuntime".Work[#RootIndex].Payload.Records[#Slot].WriteKey := "FRK_ConfigScratch".Entry.WriteKey;
        "FRK_SetRuntime".Work[#RootIndex].Payload.Records[#Slot].Revision := "FRK_ConfigScratch".Entry.WriteRevision;
        "FRK_SetRuntime".Work[#RootIndex].Payload.Records[#Slot].Kind := "FRK_ConfigScratch".Entry.ConfigKind;
        "FRK_SetRuntime".Work[#RootIndex].Payload.Records[#Slot].ValueType := "FRK_ConfigScratch".Entry.ValueType;
        "FRK_SetRuntime".Work[#RootIndex].Payload.Records[#Slot].ValueText := WSTRING_TO_STRING("FRK_ConfigScratch".Entry.ValueText);
        "FRK_SetRuntime".Work[#RootIndex].Payload.Info.RecordCount := #Slot;
    ELSE
        #Slot := "FRK_SetCheck"(RootIndex := #RootIndex, Scope := #Scope, Access := #Access, Ready := #Ready AND (#Phase = 4 OR "FRK_Line".Ready), WriteAccess := #Phase <> 3, ReserveTarget := FALSE);
        IF #Slot = 0 THEN RETURN; END_IF;
        IF #Phase = 1 OR #Phase = 4 THEN
    "FRK_LineSetStage".Values.ShiftActiveDays[3] := LINT_TO_DINT("FRK_ConfigScratch".Value.Number);
        END_IF;
    END_IF;
    "FRK_LineDef"(FieldIndex := 21);
    "FRK_SetRuntime".Work[#RootIndex].RejectScope := #Scope; "FRK_SetRuntime".Work[#RootIndex].RejectKey := "FRK_ConfigScratch".Entry.WriteKey;
    IF #Phase = 0 OR #Phase = 5 THEN
        IF #Phase = 5 AND NOT "FRK_ConfigDataAllowed"(Access := #Access, ForWrite := FALSE, Scope := #Scope) THEN RETURN; END_IF;
        "FRK_LineValue"(FieldIndex := 21, Values := "FRK_Line".Data.Values);
        IF NOT "FRK_ConfigValidate"(Text := "FRK_ConfigScratch".Entry.ValueText)
            OR "FRK_SetRuntime".Work[#RootIndex].Payload.Info.RecordCount >= 29 THEN RETURN; END_IF;
        #Slot := "FRK_SetRuntime".Work[#RootIndex].Payload.Info.RecordCount + 1;
        "FRK_SetRuntime".Work[#RootIndex].Payload.Records[#Slot].Scope := #Scope;
        "FRK_SetRuntime".Work[#RootIndex].Payload.Records[#Slot].WriteKey := "FRK_ConfigScratch".Entry.WriteKey;
        "FRK_SetRuntime".Work[#RootIndex].Payload.Records[#Slot].Revision := "FRK_ConfigScratch".Entry.WriteRevision;
        "FRK_SetRuntime".Work[#RootIndex].Payload.Records[#Slot].Kind := "FRK_ConfigScratch".Entry.ConfigKind;
        "FRK_SetRuntime".Work[#RootIndex].Payload.Records[#Slot].ValueType := "FRK_ConfigScratch".Entry.ValueType;
        "FRK_SetRuntime".Work[#RootIndex].Payload.Records[#Slot].ValueText := WSTRING_TO_STRING("FRK_ConfigScratch".Entry.ValueText);
        "FRK_SetRuntime".Work[#RootIndex].Payload.Info.RecordCount := #Slot;
    ELSE
        #Slot := "FRK_SetCheck"(RootIndex := #RootIndex, Scope := #Scope, Access := #Access, Ready := #Ready AND (#Phase = 4 OR "FRK_Line".Ready), WriteAccess := #Phase <> 3, ReserveTarget := FALSE);
        IF #Slot = 0 THEN RETURN; END_IF;
        IF #Phase = 1 OR #Phase = 4 THEN
    "FRK_LineSetStage".Values.ShiftTarget[3] := LINT_TO_DINT("FRK_ConfigScratch".Value.Number);
        END_IF;
    END_IF;
    "FRK_LineDef"(FieldIndex := 22);
    "FRK_SetRuntime".Work[#RootIndex].RejectScope := #Scope; "FRK_SetRuntime".Work[#RootIndex].RejectKey := "FRK_ConfigScratch".Entry.WriteKey;
    IF #Phase = 0 OR #Phase = 5 THEN
        IF #Phase = 5 AND NOT "FRK_ConfigDataAllowed"(Access := #Access, ForWrite := FALSE, Scope := #Scope) THEN RETURN; END_IF;
        "FRK_LineValue"(FieldIndex := 22, Values := "FRK_Line".Data.Values);
        IF NOT "FRK_ConfigValidate"(Text := "FRK_ConfigScratch".Entry.ValueText)
            OR "FRK_SetRuntime".Work[#RootIndex].Payload.Info.RecordCount >= 29 THEN RETURN; END_IF;
        #Slot := "FRK_SetRuntime".Work[#RootIndex].Payload.Info.RecordCount + 1;
        "FRK_SetRuntime".Work[#RootIndex].Payload.Records[#Slot].Scope := #Scope;
        "FRK_SetRuntime".Work[#RootIndex].Payload.Records[#Slot].WriteKey := "FRK_ConfigScratch".Entry.WriteKey;
        "FRK_SetRuntime".Work[#RootIndex].Payload.Records[#Slot].Revision := "FRK_ConfigScratch".Entry.WriteRevision;
        "FRK_SetRuntime".Work[#RootIndex].Payload.Records[#Slot].Kind := "FRK_ConfigScratch".Entry.ConfigKind;
        "FRK_SetRuntime".Work[#RootIndex].Payload.Records[#Slot].ValueType := "FRK_ConfigScratch".Entry.ValueType;
        "FRK_SetRuntime".Work[#RootIndex].Payload.Records[#Slot].ValueText := WSTRING_TO_STRING("FRK_ConfigScratch".Entry.ValueText);
        "FRK_SetRuntime".Work[#RootIndex].Payload.Info.RecordCount := #Slot;
    ELSE
        #Slot := "FRK_SetCheck"(RootIndex := #RootIndex, Scope := #Scope, Access := #Access, Ready := #Ready AND (#Phase = 4 OR "FRK_Line".Ready), WriteAccess := #Phase <> 3, ReserveTarget := FALSE);
        IF #Slot = 0 THEN RETURN; END_IF;
        IF #Phase = 1 OR #Phase = 4 THEN
    "FRK_LineSetStage".Values.ShiftStartMin[4] := LINT_TO_DINT("FRK_ConfigScratch".Value.Number);
        END_IF;
    END_IF;
    "FRK_LineDef"(FieldIndex := 23);
    "FRK_SetRuntime".Work[#RootIndex].RejectScope := #Scope; "FRK_SetRuntime".Work[#RootIndex].RejectKey := "FRK_ConfigScratch".Entry.WriteKey;
    IF #Phase = 0 OR #Phase = 5 THEN
        IF #Phase = 5 AND NOT "FRK_ConfigDataAllowed"(Access := #Access, ForWrite := FALSE, Scope := #Scope) THEN RETURN; END_IF;
        "FRK_LineValue"(FieldIndex := 23, Values := "FRK_Line".Data.Values);
        IF NOT "FRK_ConfigValidate"(Text := "FRK_ConfigScratch".Entry.ValueText)
            OR "FRK_SetRuntime".Work[#RootIndex].Payload.Info.RecordCount >= 29 THEN RETURN; END_IF;
        #Slot := "FRK_SetRuntime".Work[#RootIndex].Payload.Info.RecordCount + 1;
        "FRK_SetRuntime".Work[#RootIndex].Payload.Records[#Slot].Scope := #Scope;
        "FRK_SetRuntime".Work[#RootIndex].Payload.Records[#Slot].WriteKey := "FRK_ConfigScratch".Entry.WriteKey;
        "FRK_SetRuntime".Work[#RootIndex].Payload.Records[#Slot].Revision := "FRK_ConfigScratch".Entry.WriteRevision;
        "FRK_SetRuntime".Work[#RootIndex].Payload.Records[#Slot].Kind := "FRK_ConfigScratch".Entry.ConfigKind;
        "FRK_SetRuntime".Work[#RootIndex].Payload.Records[#Slot].ValueType := "FRK_ConfigScratch".Entry.ValueType;
        "FRK_SetRuntime".Work[#RootIndex].Payload.Records[#Slot].ValueText := WSTRING_TO_STRING("FRK_ConfigScratch".Entry.ValueText);
        "FRK_SetRuntime".Work[#RootIndex].Payload.Info.RecordCount := #Slot;
    ELSE
        #Slot := "FRK_SetCheck"(RootIndex := #RootIndex, Scope := #Scope, Access := #Access, Ready := #Ready AND (#Phase = 4 OR "FRK_Line".Ready), WriteAccess := #Phase <> 3, ReserveTarget := FALSE);
        IF #Slot = 0 THEN RETURN; END_IF;
        IF #Phase = 1 OR #Phase = 4 THEN
    "FRK_LineSetStage".Values.ShiftDurationMin[4] := LINT_TO_DINT("FRK_ConfigScratch".Value.Number);
        END_IF;
    END_IF;
    "FRK_LineDef"(FieldIndex := 24);
    "FRK_SetRuntime".Work[#RootIndex].RejectScope := #Scope; "FRK_SetRuntime".Work[#RootIndex].RejectKey := "FRK_ConfigScratch".Entry.WriteKey;
    IF #Phase = 0 OR #Phase = 5 THEN
        IF #Phase = 5 AND NOT "FRK_ConfigDataAllowed"(Access := #Access, ForWrite := FALSE, Scope := #Scope) THEN RETURN; END_IF;
        "FRK_LineValue"(FieldIndex := 24, Values := "FRK_Line".Data.Values);
        IF NOT "FRK_ConfigValidate"(Text := "FRK_ConfigScratch".Entry.ValueText)
            OR "FRK_SetRuntime".Work[#RootIndex].Payload.Info.RecordCount >= 29 THEN RETURN; END_IF;
        #Slot := "FRK_SetRuntime".Work[#RootIndex].Payload.Info.RecordCount + 1;
        "FRK_SetRuntime".Work[#RootIndex].Payload.Records[#Slot].Scope := #Scope;
        "FRK_SetRuntime".Work[#RootIndex].Payload.Records[#Slot].WriteKey := "FRK_ConfigScratch".Entry.WriteKey;
        "FRK_SetRuntime".Work[#RootIndex].Payload.Records[#Slot].Revision := "FRK_ConfigScratch".Entry.WriteRevision;
        "FRK_SetRuntime".Work[#RootIndex].Payload.Records[#Slot].Kind := "FRK_ConfigScratch".Entry.ConfigKind;
        "FRK_SetRuntime".Work[#RootIndex].Payload.Records[#Slot].ValueType := "FRK_ConfigScratch".Entry.ValueType;
        "FRK_SetRuntime".Work[#RootIndex].Payload.Records[#Slot].ValueText := WSTRING_TO_STRING("FRK_ConfigScratch".Entry.ValueText);
        "FRK_SetRuntime".Work[#RootIndex].Payload.Info.RecordCount := #Slot;
    ELSE
        #Slot := "FRK_SetCheck"(RootIndex := #RootIndex, Scope := #Scope, Access := #Access, Ready := #Ready AND (#Phase = 4 OR "FRK_Line".Ready), WriteAccess := #Phase <> 3, ReserveTarget := FALSE);
        IF #Slot = 0 THEN RETURN; END_IF;
        IF #Phase = 1 OR #Phase = 4 THEN
    "FRK_LineSetStage".Values.ShiftActiveDays[4] := LINT_TO_DINT("FRK_ConfigScratch".Value.Number);
        END_IF;
    END_IF;
    "FRK_LineDef"(FieldIndex := 25);
    "FRK_SetRuntime".Work[#RootIndex].RejectScope := #Scope; "FRK_SetRuntime".Work[#RootIndex].RejectKey := "FRK_ConfigScratch".Entry.WriteKey;
    IF #Phase = 0 OR #Phase = 5 THEN
        IF #Phase = 5 AND NOT "FRK_ConfigDataAllowed"(Access := #Access, ForWrite := FALSE, Scope := #Scope) THEN RETURN; END_IF;
        "FRK_LineValue"(FieldIndex := 25, Values := "FRK_Line".Data.Values);
        IF NOT "FRK_ConfigValidate"(Text := "FRK_ConfigScratch".Entry.ValueText)
            OR "FRK_SetRuntime".Work[#RootIndex].Payload.Info.RecordCount >= 29 THEN RETURN; END_IF;
        #Slot := "FRK_SetRuntime".Work[#RootIndex].Payload.Info.RecordCount + 1;
        "FRK_SetRuntime".Work[#RootIndex].Payload.Records[#Slot].Scope := #Scope;
        "FRK_SetRuntime".Work[#RootIndex].Payload.Records[#Slot].WriteKey := "FRK_ConfigScratch".Entry.WriteKey;
        "FRK_SetRuntime".Work[#RootIndex].Payload.Records[#Slot].Revision := "FRK_ConfigScratch".Entry.WriteRevision;
        "FRK_SetRuntime".Work[#RootIndex].Payload.Records[#Slot].Kind := "FRK_ConfigScratch".Entry.ConfigKind;
        "FRK_SetRuntime".Work[#RootIndex].Payload.Records[#Slot].ValueType := "FRK_ConfigScratch".Entry.ValueType;
        "FRK_SetRuntime".Work[#RootIndex].Payload.Records[#Slot].ValueText := WSTRING_TO_STRING("FRK_ConfigScratch".Entry.ValueText);
        "FRK_SetRuntime".Work[#RootIndex].Payload.Info.RecordCount := #Slot;
    ELSE
        #Slot := "FRK_SetCheck"(RootIndex := #RootIndex, Scope := #Scope, Access := #Access, Ready := #Ready AND (#Phase = 4 OR "FRK_Line".Ready), WriteAccess := #Phase <> 3, ReserveTarget := FALSE);
        IF #Slot = 0 THEN RETURN; END_IF;
        IF #Phase = 1 OR #Phase = 4 THEN
    "FRK_LineSetStage".Values.ShiftTarget[4] := LINT_TO_DINT("FRK_ConfigScratch".Value.Number);
        END_IF;
    END_IF;
    "FRK_LineDef"(FieldIndex := 26);
    "FRK_SetRuntime".Work[#RootIndex].RejectScope := #Scope; "FRK_SetRuntime".Work[#RootIndex].RejectKey := "FRK_ConfigScratch".Entry.WriteKey;
    IF #Phase = 0 OR #Phase = 5 THEN
        IF #Phase = 5 AND NOT "FRK_ConfigDataAllowed"(Access := #Access, ForWrite := FALSE, Scope := #Scope) THEN RETURN; END_IF;
        "FRK_LineValue"(FieldIndex := 26, Values := "FRK_Line".Data.Values);
        IF NOT "FRK_ConfigValidate"(Text := "FRK_ConfigScratch".Entry.ValueText)
            OR "FRK_SetRuntime".Work[#RootIndex].Payload.Info.RecordCount >= 29 THEN RETURN; END_IF;
        #Slot := "FRK_SetRuntime".Work[#RootIndex].Payload.Info.RecordCount + 1;
        "FRK_SetRuntime".Work[#RootIndex].Payload.Records[#Slot].Scope := #Scope;
        "FRK_SetRuntime".Work[#RootIndex].Payload.Records[#Slot].WriteKey := "FRK_ConfigScratch".Entry.WriteKey;
        "FRK_SetRuntime".Work[#RootIndex].Payload.Records[#Slot].Revision := "FRK_ConfigScratch".Entry.WriteRevision;
        "FRK_SetRuntime".Work[#RootIndex].Payload.Records[#Slot].Kind := "FRK_ConfigScratch".Entry.ConfigKind;
        "FRK_SetRuntime".Work[#RootIndex].Payload.Records[#Slot].ValueType := "FRK_ConfigScratch".Entry.ValueType;
        "FRK_SetRuntime".Work[#RootIndex].Payload.Records[#Slot].ValueText := WSTRING_TO_STRING("FRK_ConfigScratch".Entry.ValueText);
        "FRK_SetRuntime".Work[#RootIndex].Payload.Info.RecordCount := #Slot;
    ELSE
        #Slot := "FRK_SetCheck"(RootIndex := #RootIndex, Scope := #Scope, Access := #Access, Ready := #Ready AND (#Phase = 4 OR "FRK_Line".Ready), WriteAccess := #Phase <> 3, ReserveTarget := FALSE);
        IF #Slot = 0 THEN RETURN; END_IF;
        IF #Phase = 1 OR #Phase = 4 THEN
    "FRK_LineSetStage".Values.ShiftStartMin[5] := LINT_TO_DINT("FRK_ConfigScratch".Value.Number);
        END_IF;
    END_IF;
    "FRK_LineDef"(FieldIndex := 27);
    "FRK_SetRuntime".Work[#RootIndex].RejectScope := #Scope; "FRK_SetRuntime".Work[#RootIndex].RejectKey := "FRK_ConfigScratch".Entry.WriteKey;
    IF #Phase = 0 OR #Phase = 5 THEN
        IF #Phase = 5 AND NOT "FRK_ConfigDataAllowed"(Access := #Access, ForWrite := FALSE, Scope := #Scope) THEN RETURN; END_IF;
        "FRK_LineValue"(FieldIndex := 27, Values := "FRK_Line".Data.Values);
        IF NOT "FRK_ConfigValidate"(Text := "FRK_ConfigScratch".Entry.ValueText)
            OR "FRK_SetRuntime".Work[#RootIndex].Payload.Info.RecordCount >= 29 THEN RETURN; END_IF;
        #Slot := "FRK_SetRuntime".Work[#RootIndex].Payload.Info.RecordCount + 1;
        "FRK_SetRuntime".Work[#RootIndex].Payload.Records[#Slot].Scope := #Scope;
        "FRK_SetRuntime".Work[#RootIndex].Payload.Records[#Slot].WriteKey := "FRK_ConfigScratch".Entry.WriteKey;
        "FRK_SetRuntime".Work[#RootIndex].Payload.Records[#Slot].Revision := "FRK_ConfigScratch".Entry.WriteRevision;
        "FRK_SetRuntime".Work[#RootIndex].Payload.Records[#Slot].Kind := "FRK_ConfigScratch".Entry.ConfigKind;
        "FRK_SetRuntime".Work[#RootIndex].Payload.Records[#Slot].ValueType := "FRK_ConfigScratch".Entry.ValueType;
        "FRK_SetRuntime".Work[#RootIndex].Payload.Records[#Slot].ValueText := WSTRING_TO_STRING("FRK_ConfigScratch".Entry.ValueText);
        "FRK_SetRuntime".Work[#RootIndex].Payload.Info.RecordCount := #Slot;
    ELSE
        #Slot := "FRK_SetCheck"(RootIndex := #RootIndex, Scope := #Scope, Access := #Access, Ready := #Ready AND (#Phase = 4 OR "FRK_Line".Ready), WriteAccess := #Phase <> 3, ReserveTarget := FALSE);
        IF #Slot = 0 THEN RETURN; END_IF;
        IF #Phase = 1 OR #Phase = 4 THEN
    "FRK_LineSetStage".Values.ShiftDurationMin[5] := LINT_TO_DINT("FRK_ConfigScratch".Value.Number);
        END_IF;
    END_IF;
    "FRK_LineDef"(FieldIndex := 28);
    "FRK_SetRuntime".Work[#RootIndex].RejectScope := #Scope; "FRK_SetRuntime".Work[#RootIndex].RejectKey := "FRK_ConfigScratch".Entry.WriteKey;
    IF #Phase = 0 OR #Phase = 5 THEN
        IF #Phase = 5 AND NOT "FRK_ConfigDataAllowed"(Access := #Access, ForWrite := FALSE, Scope := #Scope) THEN RETURN; END_IF;
        "FRK_LineValue"(FieldIndex := 28, Values := "FRK_Line".Data.Values);
        IF NOT "FRK_ConfigValidate"(Text := "FRK_ConfigScratch".Entry.ValueText)
            OR "FRK_SetRuntime".Work[#RootIndex].Payload.Info.RecordCount >= 29 THEN RETURN; END_IF;
        #Slot := "FRK_SetRuntime".Work[#RootIndex].Payload.Info.RecordCount + 1;
        "FRK_SetRuntime".Work[#RootIndex].Payload.Records[#Slot].Scope := #Scope;
        "FRK_SetRuntime".Work[#RootIndex].Payload.Records[#Slot].WriteKey := "FRK_ConfigScratch".Entry.WriteKey;
        "FRK_SetRuntime".Work[#RootIndex].Payload.Records[#Slot].Revision := "FRK_ConfigScratch".Entry.WriteRevision;
        "FRK_SetRuntime".Work[#RootIndex].Payload.Records[#Slot].Kind := "FRK_ConfigScratch".Entry.ConfigKind;
        "FRK_SetRuntime".Work[#RootIndex].Payload.Records[#Slot].ValueType := "FRK_ConfigScratch".Entry.ValueType;
        "FRK_SetRuntime".Work[#RootIndex].Payload.Records[#Slot].ValueText := WSTRING_TO_STRING("FRK_ConfigScratch".Entry.ValueText);
        "FRK_SetRuntime".Work[#RootIndex].Payload.Info.RecordCount := #Slot;
    ELSE
        #Slot := "FRK_SetCheck"(RootIndex := #RootIndex, Scope := #Scope, Access := #Access, Ready := #Ready AND (#Phase = 4 OR "FRK_Line".Ready), WriteAccess := #Phase <> 3, ReserveTarget := FALSE);
        IF #Slot = 0 THEN RETURN; END_IF;
        IF #Phase = 1 OR #Phase = 4 THEN
    "FRK_LineSetStage".Values.ShiftActiveDays[5] := LINT_TO_DINT("FRK_ConfigScratch".Value.Number);
        END_IF;
    END_IF;
    "FRK_LineDef"(FieldIndex := 29);
    "FRK_SetRuntime".Work[#RootIndex].RejectScope := #Scope; "FRK_SetRuntime".Work[#RootIndex].RejectKey := "FRK_ConfigScratch".Entry.WriteKey;
    IF #Phase = 0 OR #Phase = 5 THEN
        IF #Phase = 5 AND NOT "FRK_ConfigDataAllowed"(Access := #Access, ForWrite := FALSE, Scope := #Scope) THEN RETURN; END_IF;
        "FRK_LineValue"(FieldIndex := 29, Values := "FRK_Line".Data.Values);
        IF NOT "FRK_ConfigValidate"(Text := "FRK_ConfigScratch".Entry.ValueText)
            OR "FRK_SetRuntime".Work[#RootIndex].Payload.Info.RecordCount >= 29 THEN RETURN; END_IF;
        #Slot := "FRK_SetRuntime".Work[#RootIndex].Payload.Info.RecordCount + 1;
        "FRK_SetRuntime".Work[#RootIndex].Payload.Records[#Slot].Scope := #Scope;
        "FRK_SetRuntime".Work[#RootIndex].Payload.Records[#Slot].WriteKey := "FRK_ConfigScratch".Entry.WriteKey;
        "FRK_SetRuntime".Work[#RootIndex].Payload.Records[#Slot].Revision := "FRK_ConfigScratch".Entry.WriteRevision;
        "FRK_SetRuntime".Work[#RootIndex].Payload.Records[#Slot].Kind := "FRK_ConfigScratch".Entry.ConfigKind;
        "FRK_SetRuntime".Work[#RootIndex].Payload.Records[#Slot].ValueType := "FRK_ConfigScratch".Entry.ValueType;
        "FRK_SetRuntime".Work[#RootIndex].Payload.Records[#Slot].ValueText := WSTRING_TO_STRING("FRK_ConfigScratch".Entry.ValueText);
        "FRK_SetRuntime".Work[#RootIndex].Payload.Info.RecordCount := #Slot;
    ELSE
        #Slot := "FRK_SetCheck"(RootIndex := #RootIndex, Scope := #Scope, Access := #Access, Ready := #Ready AND (#Phase = 4 OR "FRK_Line".Ready), WriteAccess := #Phase <> 3, ReserveTarget := FALSE);
        IF #Slot = 0 THEN RETURN; END_IF;
        IF #Phase = 1 OR #Phase = 4 THEN
    "FRK_LineSetStage".Values.ShiftTarget[5] := LINT_TO_DINT("FRK_ConfigScratch".Value.Number);
        END_IF;
    END_IF;
    IF (#Phase = 1 OR #Phase = 4) AND NOT "FRK_LineValid"(Values := "FRK_LineSetStage".Values) THEN RETURN; END_IF;
    #FRK_LineSetWalk := TRUE;
END_FUNCTION
